// SIMATIC STEP 7 (V5.x) project ex14
// CPU: CPU 314
// station: Matériel
// station: SIMATIC 300(1)
// station: P_ADR_BUS
// program: Programme S7(1)

SYMBOL_TABLE
"SCALE"	FC 105	FC 105	// Scaling Values
"UNSCALE"	FC 106	FC 106	// Unscaling Values
"ROUGE"	Q 0.0	BOOL
"VERT"	Q 0.1	BOOL
"FOUR"	Q 0.2	BOOL
END_SYMBOL_TABLE

// FC 105: know-how protected block, not included

// FC 106: know-how protected block, not included

ORGANIZATION_BLOCK OB 1
TITLE = "Main Program Sweep (Cycle)"
VERSION : 0.1
VAR_TEMP
  OB1_EV_CLASS : BYTE ;	//Bits 0-3 = 1 (Coming event), Bits 4-7 = 1 (Event class 1)
  OB1_SCAN_1 : BYTE ;	//1 (Cold restart scan 1 of OB 1), 3 (Scan 2-n of OB 1)
  OB1_PRIORITY : BYTE ;	//Priority of OB Execution
  OB1_OB_NUMBR : BYTE ;	//1 (Organization block 1, OB1)
  OB1_RESERVED_1 : BYTE ;	//Reserved for system
  OB1_RESERVED_2 : BYTE ;	//Reserved for system
  OB1_PREV_CYCLE : INT ;	//Cycle time of previous OB1 scan (milliseconds)
  OB1_MIN_CYCLE : INT ;	//Minimum cycle time of OB1 (milliseconds)
  OB1_MAX_CYCLE : INT ;	//Maximum cycle time of OB1 (milliseconds)
  OB1_DATE_TIME : DATE_AND_TIME ;	//Date and time OB1 started
END_VAR
BEGIN
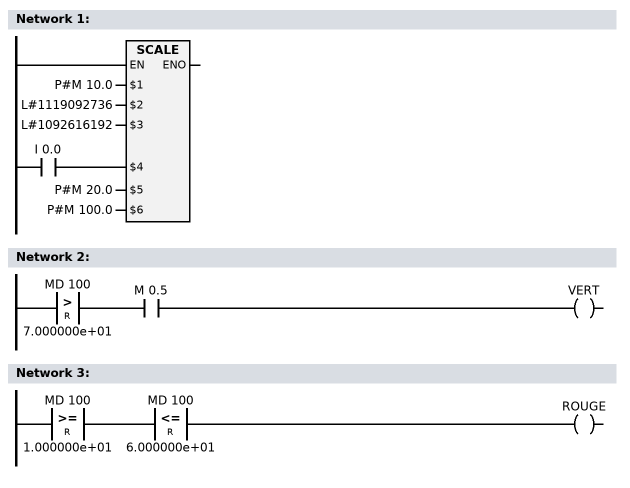
NETWORK
TITLE =
      A     I 0.0;
      =     L 20.0;
      BLD   103;
      CALL  "SCALE" (
           $1                       := P#M 10.0,
           $2                       := L#1119092736,
           $3                       := L#1092616192,
           $4                       := L 20.0,
           $5                       := P#M 20.0,
           $6                       := P#M 100.0);
      NOP   0;
NETWORK
TITLE =
      A(;
      L     MD 100;
      L     7.000000e+01;
      >R;
      );
      A     M 0.5;
      =     "VERT";
NETWORK
TITLE =
      A(;
      L     MD 100;
      L     1.000000e+01;
      >=R;
      );
      A(;
      L     MD 100;
      L     6.000000e+01;
      <=R;
      );
      =     "ROUGE";
END_ORGANIZATION_BLOCK
